(* IEC 61131-3 sources: plcassist-cli/packages/volt-lsp-iec/test-corpus/pro2193/Device/Plc Logic/Application/09 Misc/Library Manager/CmpChecksum, 7 files *)

(* ---- CRC16FINISH.fun ---- *)
FUNCTION CRC16FINISH : WORD
VAR_INPUT
	ULCRC : WORD;
END_VAR
END_FUNCTION

(* ---- CRC16INIT.fun ---- *)
FUNCTION CRC16INIT : WORD
END_FUNCTION

(* ---- CRC16UPDATE.fun ---- *)
FUNCTION CRC16UPDATE : WORD
VAR_INPUT
	ULCRC : WORD;
	PDATA : POINTER TO BYTE;
	ULSIZE : __XWORD;
END_VAR
END_FUNCTION

(* ---- CRC32FINISH.fun ---- *)
FUNCTION CRC32FINISH : DWORD
VAR_INPUT
	ULCRC : DWORD;
END_VAR
END_FUNCTION

(* ---- CRC32INIT.fun ---- *)
FUNCTION CRC32INIT : DWORD
END_FUNCTION

(* ---- CRC32UPDATE.fun ---- *)
FUNCTION CRC32UPDATE : DWORD
VAR_INPUT
	ULCRC : DWORD;
	PDATA : POINTER TO BYTE;
	ULSIZE : __XWORD;
END_VAR
END_FUNCTION

(* ---- CRC32UPDATE2.fun ---- *)
FUNCTION CRC32UPDATE2 : DWORD
VAR_INPUT
	ULCRC : DWORD;
	PDATA : POINTER TO BYTE;
	ULSIZE : __XWORD;
END_VAR
END_FUNCTION
